(* IEC 61131-3 sources: st-analyze/src/plc/workspace, 15 files *)

(* ---- alias1.st ---- *)
TYPE
	China: STRUCT
	 provinceId, qw, iuy, bb: STRING;
	 province: Province;
	 a: INT;
   END_STRUCT
END_TYPE

(* ---- china.st ---- *)
TYPE
	China: STRUCT
	 provinceId,qw,iuy,bb: INT;
	 province: Province;
	 a: CTU;
   END_STRUCT
END_TYPE

(* ---- city.st ---- *)
TYPE
	City: STRUCT
	 cityId33: INT;
	 region: Region;
	 dtTimeNow666: DATE_AND_TIME := DT#2021 - 10 - 19 - 13: 53: 00;
   END_STRUCT
END_TYPE

(* ---- province.st ---- *)
TYPE
	Province: STRUCT
	 provinceId: INT;
	 aabbcc:BOOL:=true;
	 city:City;

   END_STRUCT
END_TYPE

(* ---- region.st ---- *)
TYPE
	Region: STRUCT
	  regionName:STRING;
	  b: ARRAY [9..10] OF INT:=[1,2,3,4,5];
   END_STRUCT
END_TYPE

(* ---- union1.st ---- *)
TYPE
	TON: UNION
	 a: BOOL := FALSE;
	 b: REAL;
	 c: BOOL;

END_UNION
END_TYPE

(* ---- function1.st ---- *)
FUNCTION addNumbers: INT
VAR
    state,k : INT := 11;
    bb : INT := 22;
    sum : INT;
END_VAR
VAR_INPUT
  c:INT;
END_VAR

FOR state := 0 TO 100 BY 2 DO
  state := state + state;
  IF state >= 100 THEN
    EXIT

  END_IF
END_FOR

 RETURN state+bb;

END_FUNCTION

(* ---- function2.st ---- *)
FUNCTION addNumbers66 : INT
VAR_INPUT
    a1 : INT; // 第一个整数
    a2 : INT; // 第二个整数
    a3 : INT; // 第三个整数
    a4 : INT; // 第四个整数
END_VAR
VAR
    result : INT; // 存储中间结果
END_VAR

result := a1 + a2 + a3 + a4;
RETURN result;

END_FUNCTION

(* ---- enum1.st ---- *)
TYPE
    ColorEnum : (
        Red := 0,
        Green := 1,
        Blue := 2,
        Yellow := 3
    )
END_TYPE
  TYPE COLOR1 : (red, blue) END_TYPE
PROGRAM EnumProgram

VAR
     state: INT := 9;
     province: Province;

END_VAR
END_PROGRAM

FUNCTION_BLOCK EnumFB
VAR
     ccc,yuo: R_TRIG; // 定义一个实数类型的变量 celsius，用于存储摄氏温度
    dd: REAL:=123.89874141;
    ee:CTU;
    ff:BOOL;
    dtTimeNow:DATE_AND_TIME:=DT#2021-10-19-13:53:00;

END_VAR
END_FUNCTION_BLOCK

(* ---- functionBlock1.st ---- *)
FUNCTION_BLOCK TemperatureConverter
VAR
     ccc,mm: R_TRIG; // 定义一个实数类型的变量 celsius，用于存储摄氏温度
    dd: REAL;
    ee:LINT;
    ff:BOOL:=1;
    dtTimeNow:DATE_AND_TIME:=DT#2021-10-19-13:53:00;

END_VAR

VAR_INPUT
     aeiuqjnkjad,hh:BOOL;
	bbtrtr,ll:INT;
	cccc:STRING;
     d:INT;
END_VAR
VAR_OUTPUT
  kk:INT;
  mmty:INT;
END_VAR

VAR_EXTERNAL
    DevUniAxis1 : AXIS_REF;
END_VAR

// METHOD ConvertCelsiusToFahrenheit58(celsiusTemp: InT): REAL
// VAR
//     fahrenheitTemp: tof; // 定义一个实数类型的变量 fahrenheitTemp，用于存储转换后的华氏温度
//     celsiusTemp:REAL;

// END_VAR
// VAR_INPUT
//    ipio:STRing;

// END_VAR
//  fahrenheitTemp := celsiusTemp * 9 / 5 + 32; // 将摄氏温度转换为华氏温度

// END_METHOD

// METHOD ConvertCelsiusToFahrenheit(celsiusTemp: ReAL): REAL
// VAR
//     fahrenheitTemp: REAL; // 定义一个实数类型的变量 fahrenheitTemp，用于存储转换后的华氏温度
//     celsiusTemp:REAL;
// END_VAR
//  fahrenheitTemp := celsiusTemp * 9 / 5 + 32; // 将摄氏温度转换为华氏温度

// END_METHOD

END_FUNCTION_BLOCK

(* ---- functionBlock2.st ---- *)
FUNCTION_BLOCK TemperatureConverter2
VAR
     ccc: R_TRIG; // 定义一个实数类型的变量 celsius，用于存储摄氏温度
    dd, mn, kk, hh: REAL;
    ee, hj, qwer: LINT;
    ff, zx, jj, as, rr: China;
    dt, pp, ii: DATE_AND_TIME := DT#2021 - 10 - 19 - 13: 53: 00;

END_VAR

// METHOD ConvertCelsiusToFahrenheit365(celsiusTemp: REAL): REAL
// VAR
// fahrenheitTemp: R_TRIG; // 定义一个实数类型的变量 fahrenheitTemp，用于存储转换后的华氏温度
// region: DINT;
// END_VAR
// VAR_INPUT
// ipio: STRING;
// END_VAR
// fahrenheitTemp := celsiusTemp * 9 / 5 + 32; // 将摄氏温度转换为华氏温度

// END_METHOD

METHOD ConvertCelsiusToFahrenheit6(celsiusTemp: REAL): REAL
VAR
fahrenheitTemp: REAL; // 定义一个实数类型的变量 fahrenheitTemp，用于存储转换后的华氏温度
celsiusTemp: REAL;
END_VAR
 // 将摄氏温度转换为华氏温度

 END_METHOD

ee:=12;
END_FUNCTION_BLOCK

(* ---- main.st ---- *)
// TYPE
// 	China: STRUCT
// 	 provinceId, qw, iuy, bb: INT;
// 	 province: Province;
// 	 a: CTU;
// END_STRUCT
// END_TYPE

PROGRAM Test
VAR
	a: AXIS_REF;
	b: SMC_TrackAxis;
    c: SMC_TP;
	d: TON;
	mode: RunMode;
	libEnum: MC_BUFFER_MODE;
	e: Province;
	f: MC_Direction;
	g: China;
	h:INT;
	aa:sint;
END_VAR
VAR_IN_OUT
	Variable: BOOL; (* Comment *)
END_VAR

VAR_EXTERNAL
    gStart : BOOL;
    gCount : INT;
    gLamp  : BOOL;
	aa:TON;
END_VAR

IF GVL.gStart THEN
    GVL.gCount := GVL.gCount + 1;
END_IF;

IF GVL_1.aa.Q THEN
    GVL.gCount := GVL.gCount + 1;
END_IF;

mode := RunMode#MANUAL;
libEnum := MC_BUFFER_MODE#Aborting;
c.delta_time := T#3h2m33s11ms;
d.IN := 1;
e.city.region.regionName := 'Beijing';
f := MC_Direction#fastest;

e.city.cityId33:=123;
h:=-90;

aa:=0;

END_PROGRAM

(* ---- program2.st ---- *)
PROGRAM PLC_PRG
VAR
     state: INT;
     result: INT := 19999;
    result2: STRING := 'qw';
    china,china2: China;
    a: WORD := 65137;
    voltage: REAL := 1235.754289;
    tempConverter: TemperatureConverter2;
    t, o: TIME_OF_DAY;
    b: ARRAY [9..10] OF INT := [1, 0, 1, 1, 1];
    tHold: TIME:= T#3h2m33s11ms;
    dteStart: DATE:= DATE#2020-10-19;
    dtTimeNow: DATE_AND_TIME:= DT#2021-10-19-13:53:00;
    todTimer: TIME_OF_DAY:= TOD#08:08:59.555;
    t33:TON;
    testDateTime:DT:=DT#2024-04-16-23:33:00.22;
	testTod:TOD:=TOD#23:33:00.22;
    // o: DATE :=DATE#2021-10-19;
END_VAR

tempConverter.dd:=12.34;
 //voltage := tempConverter.ConvertCelsiusToFahrenheit365(12.357778); // 将摄氏温度转换为华氏温度
 china.province.city.region.regionName := '小店区';
// result := addNumbers(5, 7,8,9);
CASE state OF
1, 3, 5, 7, 8, 10, 12:
state := 12;
15..100:
state := 15;
ELSE
state := 18;
END_CASE

IF state > 10 THEN
state := 1 / 3;
ELSIF state > result THEN
state := state;
ELSE
state := 3;
END_IF

REPEAT
state := state + 1; // 每次循环计数器加1
// 在这里可以添加其他逻辑操作

UNTIL state >= 5 // 当计数器达到5时结束循环
END_REPEAT

WHILE a <> 0 DO
  b := b * 2;
  a := a - 1;
END_WHILE
FOR  state:= 0  TO 100 BY 2 DO
  state:=5+state;
  IF state>=100 THEN
    EXIT
  END_IF
END_FOR

END_PROGRAM

(* ---- test33.st ---- *)
PROGRAM Test1155667788
VAR
	a: BOOL;
	c: BOOL;
	d: BOOL;
	e: INT;
	qww: INT;
	g: INT;
	b: CTU;
	dd:USINT:=0;
	asd:SEMA;
	mmm:CTU_DINT;
END_VAR

(* generate 【segmentId 174237778419740866】 code start *)
IF a THEN
 CTU(CU := c, R := d, PV := e, Q => c, CV => g);
END_IF
(* generate 【segmentId 174237778419740866】 code end *)

END_PROGRAM

(* ---- ton.st ---- *)
PROGRAM Test
VAR
	a: BOOL;
	b: BOOL;
	c: BOOL;
	f: BOOL;
	h: BOOL;
	i: BOOL;
	g: BOOL;
	p: BOOL;
	e: BOOL;
	d: SR;
	k: BOOL;
	l: BOOL;
	m: INT;
	n: BOOL;
	o: INT;
	j: CTU;
	bb:BOOL;
END_VAR

(* generate 【segmentId 174556890774562716】 code start *)
d(S1 := a, R := e, Q1 => );
IF ((a AND ((b AND c) OR i OR (g AND h AND f))) OR ((d.Q1 AND f))) THEN
 CTU(CU := k, R := l, PV := m, Q => n, CV => o);
END_IF
IF (a AND ((b AND c) OR i OR (g AND h AND f))) OR ((d.Q1 AND f)) THEN
 p := TRUE;
END_IF
(* generate 【segmentId 174556890774562716】 code end *)

END_PROGRAM
